// TIA Portal V21 export
FUNCTION_BLOCK "Guard"   // FB5, F_FBD
{ S7_Optimized_Access := 'TRUE' }
// A guard door: open while its switch is not closed.
   VAR_INPUT
      closed : Bool;
   END_VAR
   VAR_OUTPUT
      open : Bool;
   END_VAR
BEGIN

REGION Network 1: Open guard
   // The guard is open while its switch is not closed.
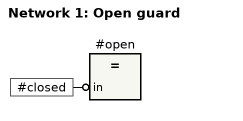
   #open := NOT #closed;
END_REGION
END_FUNCTION_BLOCK
